// TIA Portal V20 export
Screen "MB190RB06 LOADING STAND FIFO"  1276x673
  ScreenItem "线_1" at 0,65 size 1362x0  Type=HmiLine
  ScreenItem "permanentareaborderrectangle" at 0,0 size 0x0  Type=HmiRectangle
  ScreenItem "Button_Back" at 2,2 size 90x47  Type=HmiButton
  ScreenItem "OPMode4_Foreground_Blocked" at 1160,0 size 88x58  Type=HmiGraphicView
  ScreenItem "面板容器_2" at 1160,0 size 88x58  Type=HmiFaceplateContainer
  ScreenItem "Title_OPOverview_ScreenOverview_X390_Y2" at 433,13 size 500x30  Type=HmiTextBox
  ScreenItem "Faceplate container_1" at 11,65 size 1240x580  Type=HmiFaceplateContainer
